PROGRAM prg_TriBlender
VAR
	enumCurrentState	: ENUM_CurrentState;
	FB_SetProductionParams:FB_SetProductionParams;
//stTriBlender		: ST_TriBlender;
	
	sStateDescription		: STRING;
	sStateInstructions		: STRING;
	iCirculationTimeLeft	: UINT;
	bContinue				: BOOL;
	iCurrentMixingComponent	: INT;
	
	tonStageCirculation		: TON;
	
	///For Visu
	bDisableTime			: BOOL;
	bDisableAmount			: BOOL;
	bDisableName			: BOOL;
	bDisableButton			: BOOL;
	wButtonColor			: DWORD;
	
	trig_JumpToCirScreen	: R_TRIG;

	i						: INT;
	bTesting: BOOL;
END_VAR
VAR_IN_OUT
	stTriblender			: ST_TriBlender;
	fb_TriBlenderPump		: FB_Pump;
END_VAR
VAR_INPUT
	arrComponents	: ARRAY [0..g_Prod.cMaxCompInProduct-1] OF ST_Component;
END_VAR

trig_JumpToCirScreen(CLK:= stTriblender.bStartDisolving);

IF trig_JumpToCirScreen.Q THEN
	VisuElems.CurrentVisu:= 'Main';	
END_IF

Init_act_MixingStates();

stTriblender.bPumpOnFdbk:= fb_TriBlenderPump.bRun;

FB_SetProductionParams(stProdParams:=g_Data.arr_ProdTank[0],bTankInProduction:=bTesting,iActualWaterAmount:=100,stTriBlender:=g_Data.stTriBlender);

ACTION CheckIfLast_entry:
bDisableButton:=FALSE;

fb_TriBlenderPump.m_Stop();
bContinue:=FALSE;
END_ACTION

ACTION FlowOrPressureError_entry:
stTriblender.bError:=TRUE;
stTriblender.sErrorDescription:='Pressure or flow error';
VisuElems.CurrentVisu:= 'StartVisu';
END_ACTION

ACTION Init_act_MixingStates:
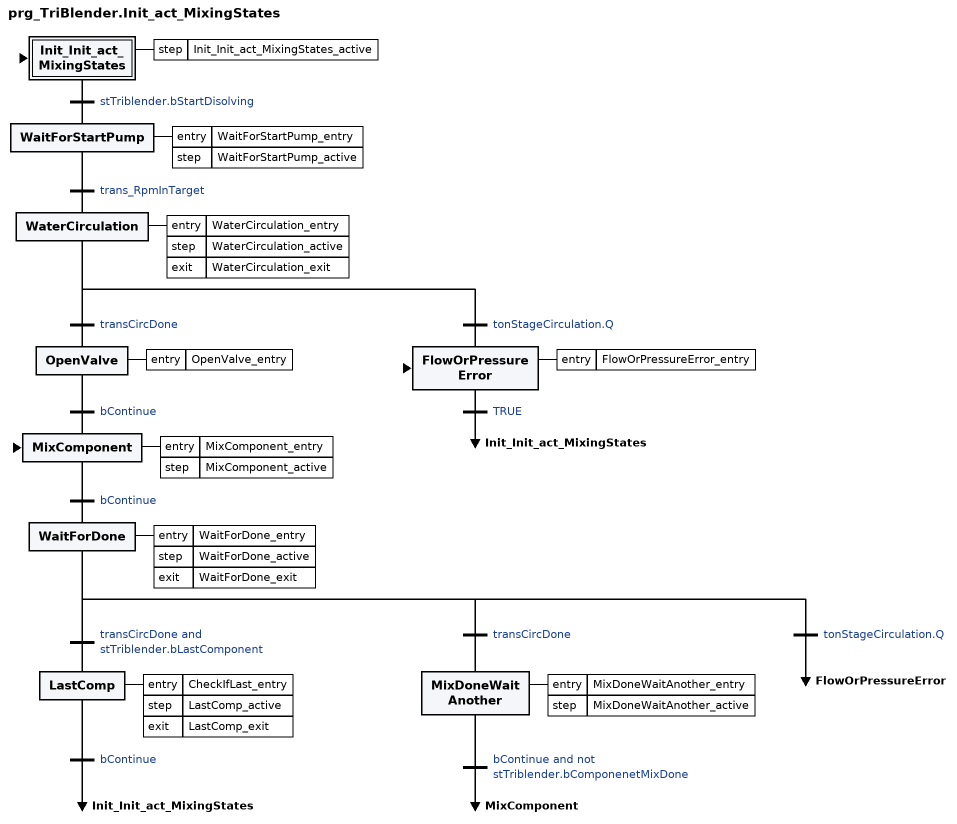
INITIAL_STEP Init_Init_act_MixingStates:
    Init_Init_act_MixingStates_active(N);  // step action
END_STEP
TRANSITION FROM Init_Init_act_MixingStates TO WaitForStartPump
    := stTriblender.bStartDisolving;
END_TRANSITION
STEP WaitForStartPump:
    WaitForStartPump_entry(P1);  // entry action
    WaitForStartPump_active(N);  // step action
END_STEP
TRANSITION FROM WaitForStartPump TO WaterCirculation
    := trans_RpmInTarget;
END_TRANSITION
STEP WaterCirculation:
    WaterCirculation_entry(P1);  // entry action
    WaterCirculation_active(N);  // step action
    WaterCirculation_exit(P0);  // exit action
END_STEP
TRANSITION FROM WaterCirculation TO OpenValve
    := transCircDone;
END_TRANSITION
TRANSITION FROM WaterCirculation TO FlowOrPressureError
    := tonStageCirculation.Q;
END_TRANSITION
STEP FlowOrPressureError:
    FlowOrPressureError_entry(P1);  // entry action
END_STEP
TRANSITION FROM FlowOrPressureError TO Init_Init_act_MixingStates
    := TRUE;
END_TRANSITION
STEP OpenValve:
    OpenValve_entry(P1);  // entry action
END_STEP
TRANSITION FROM OpenValve TO MixComponent
    := bContinue;
END_TRANSITION
STEP MixComponent:
    MixComponent_entry(P1);  // entry action
    MixComponent_active(N);  // step action
END_STEP
TRANSITION FROM MixComponent TO WaitForDone
    := bContinue;
END_TRANSITION
STEP WaitForDone:
    WaitForDone_entry(P1);  // entry action
    WaitForDone_active(N);  // step action
    WaitForDone_exit(P0);  // exit action
END_STEP
TRANSITION FROM WaitForDone TO LastComp
    := transCircDone and stTriblender.bLastComponent;
END_TRANSITION
TRANSITION FROM WaitForDone TO MixDoneWaitAnother
    := transCircDone;
END_TRANSITION
TRANSITION FROM WaitForDone TO FlowOrPressureError
    := tonStageCirculation.Q;
END_TRANSITION
STEP MixDoneWaitAnother:
    MixDoneWaitAnother_entry(P1);  // entry action
    MixDoneWaitAnother_active(N);  // step action
END_STEP
TRANSITION FROM MixDoneWaitAnother TO MixComponent
    := bContinue and not stTriblender.bComponenetMixDone;
END_TRANSITION
STEP LastComp:
    CheckIfLast_entry(P1);  // entry action
    LastComp_active(N);  // step action
    LastComp_exit(P0);  // exit action
END_STEP
TRANSITION FROM LastComp TO Init_Init_act_MixingStates
    := bContinue;
END_TRANSITION
// branch label Branch1_Init_act_MixingStates
// branch label Branch2_Init_act_MixingStates
// branch label Branch0_Init_act_MixingStates
END_ACTION

ACTION Init_Init_act_MixingStates_active:
sStateDescription	:='Triblender valve closed';
sStateInstructions	:= 'Close triblender valve';

bDisableAmount:=TRUE;
bDisableName:=TRUE;
bDisableTime:=TRUE;

wButtonColor:=16#FFC0C0C0;
stTriblender.bError:=FALSE;
stTriblender.bDisolvingDone:=FALSE;
END_ACTION

ACTION LastComp_active:
wButtonColor:=16#FF00FFFF;

sStateDescription	:=	'Finish';
sStateInstructions	:= 	'LastComponentMixed';

bDisableAmount	:=FALSE;
bDisableName	:=FALSE;
bDisableTime	:=FALSE;
END_ACTION

ACTION LastComp_exit:
VisuElems.CurrentVisu:= 'StartVisu';
stTriblender.bDisolvingDone:=TRUE;
END_ACTION

ACTION MixComponent_active:
sStateDescription	:=	'Component Inside';
sStateInstructions	:= 	'Insert component in
 the specified amount';
END_ACTION

ACTION MixComponent_entry:
bContinue:=FALSE;

bDisableAmount	:=FALSE;
bDisableName	:=FALSE;
bDisableTime	:=FALSE;

wButtonColor:=16#FFFF0000;
IF iCurrentMixingComponent<g_Prod.cMaxCompInProduct-1 THEN
	stTriblender.bLastComponent:=NOT arrComponents[iCurrentMixingComponent+1].bComponentEnable;
END_IF
stTriblender.sComponenetAmount:=TO_STRING(arrComponents[iCurrentMixingComponent].rCompActWeight);
stTriblender.sComponenetName:=arrComponents[iCurrentMixingComponent].sDescription;
stTriblender.tComponenetMixingTime:=TO_TIME(arrComponents[iCurrentMixingComponent].iMixingTime*1000);
fb_TriBlenderPump.m_Run(RPM:=arrComponents[iCurrentMixingComponent].rRpmTarget);
END_ACTION

ACTION MixDoneWaitAnother_active:
sStateDescription	:='Triblender valve Opened';
sStateInstructions	:= 'Mix Component done,
 open triblender valve';
END_ACTION

ACTION MixDoneWaitAnother_entry:
bContinue:=FALSE;

bDisableAmount:=TRUE;
bDisableName:=TRUE;
bDisableTime:=TRUE;
bDisableButton:=FALSE;
VisuElems.CurrentVisu:= 'StartVisu';



wButtonColor:=16#FF00FF00;
END_ACTION

ACTION OpenValve_entry:
bContinue:=FALSE;

bDisableAmount:=TRUE;
bDisableName:=TRUE;
bDisableTime:=TRUE;
bDisableButton:=FALSE;

tonStageCirculation(IN:=FALSE);


sStateDescription	:='Triblender valve Opened';
sStateInstructions	:= 'Open triblender valve';

wButtonColor:=16#FF00FF00;
END_ACTION

TRANSITION trans_RpmInTarget:
fb_TriBlenderPump.nRPM< arrComponents[i].rRpmTarget+10 and fb_TriBlenderPump.nRPM> arrComponents[i].rRpmTarget-10
END_TRANSITION

TRANSITION transCircDone:
tonStageCirculation.Q and stTriblender.rMaxAllowedPressure> stTriblender.rPressure and stTriblender.rMinAllowedFlow< stTriblender.rFlow
END_TRANSITION

ACTION WaitForDone_active:
tonStageCirculation(IN:= TRUE,PT:=stTriblender.tComponenetMixingTime);
iCirculationTimeLeft:= TO_UINT(tonStageCirculation.PT - tonStageCirculation.ET)/1000;
bDisableButton:=TRUE;
END_ACTION

ACTION WaitForDone_entry:
wButtonColor:=16#FF0000FF;

sStateDescription	:=	'Waiting';
sStateInstructions	:= 	'Wait for mixing done';
bContinue:=FALSE;

bDisableAmount	:=FALSE;
bDisableName	:=FALSE;
bDisableTime	:=FALSE;


tonStageCirculation(IN:= FALSE);
END_ACTION

ACTION WaitForDone_exit:
stTriblender.bComponenetMixDone:=TRUE;
wButtonColor:=16#FF00FF00;

bDisableAmount	:=TRUE;
bDisableName	:=TRUE;
bDisableTime	:=TRUE;


tonStageCirculation(IN:= FALSE);
END_ACTION

ACTION WaitForStartPump_active:
sStateDescription	:='Start Water Circulation';
sStateInstructions	:= 'Start water circulation, check for leaks';
iCurrentMixingComponent:=0;
bContinue:=FALSE;
FOR i:= 0 TO g_Prod.cMaxCompInProduct-1 DO
	IF arrComponents[i].bIsWater THEN
		fb_TriBlenderPump.m_Run(RPM:=arrComponents[i].rRpmTarget);
	END_IF
END_FOR

wButtonColor:=16#FFFF0000;
END_ACTION

ACTION WaitForStartPump_entry:

stTriblender.bStartDisolving:=FALSE;
END_ACTION

ACTION WaterCirculation_active:
tonStageCirculation(IN:= stTriblender.bPumpOnFdbk,PT:=stTriblender.tWaterCirculationTimeout);
iCirculationTimeLeft:= TO_UINT(tonStageCirculation.PT - tonStageCirculation.ET)/1000;

bDisableButton:=TRUE;

sStateDescription	:='Wait for pressure and flow';
sStateInstructions	:= 'Water circulation in progress,
 check for leaks';
END_ACTION

ACTION WaterCirculation_entry:
bContinue:=FALSE;


bDisableAmount:=TRUE;
bDisableName:=TRUE;
bDisableTime:=FALSE;

tonStageCirculation(IN:=FALSE);
END_ACTION

ACTION WaterCirculation_exit:
tonStageCirculation(IN:=FALSE);
END_ACTION

END_PROGRAM

(* stored: Version 1.1.0.1, ProductVersion 3.1.4024.15
   POU prg_TriBlender: Id {9a86bf9e-8eae-4b5d-8890-d8083718f93d}, SpecialFunc None
   Folder Management: Id {c4ddd0e8-5407-4334-a94a-0f41bc69fac1}
   Action CheckIfLast_entry: Id {0ff06adb-60ce-46ea-a8ba-434fa5634d0f}
   Action FlowOrPressureError_entry: Id {35e66287-119c-40cd-b84f-fa3e256df670}
   Action Init_act_MixingStates: Id {1bb08866-a459-47a2-9078-0401e5c0bb96}
   Action Init_Init_act_MixingStates_active: Id {5b96ca2f-dac9-4416-a4c9-760e9f673ad5}
   Action LastComp_active: Id {2582a41b-802e-45c9-b5d0-7d9f66243cf9}
   Action LastComp_exit: Id {adb66592-836d-46a4-a518-d754da30efe6}
   Action MixComponent_active: Id {1cf67d45-d09f-49f5-ad87-5f9ec42fdf26}
   Action MixComponent_entry: Id {741dfb45-7e63-4493-9a19-e4aebedfdc46}
   Action MixDoneWaitAnother_active: Id {7d82f5bc-b6bc-4046-b841-839403eb7c9b}
   Action MixDoneWaitAnother_entry: Id {ef359ffe-0713-42c1-bf19-c582d7c20eb8}
   Action OpenValve_entry: Id {0d91f935-6559-426a-8a27-b3291b9477d1}
   Transition trans_RpmInTarget: Id {9c69763e-6f57-4306-994c-85c1a23b4746}
   Transition transCircDone: Id {c004dd09-02f8-4be2-a090-e7d683131b10}
   Action WaitForDone_active: Id {b01908cf-9a52-4e61-956b-d173f0b8e957}
   Action WaitForDone_entry: Id {a6f41bb9-a823-4292-995c-7ece526c63aa}
   Action WaitForDone_exit: Id {987162f7-5bc5-4025-8270-3ef2e2dd7475}
   Action WaitForStartPump_active: Id {ede2e026-6ebe-4290-b268-7d5f0ce1e1d3}
   Action WaitForStartPump_entry: Id {59115d06-ebf0-45e1-9214-3f31cd33f08b}
   Action WaterCirculation_active: Id {4f4fcdfa-6e26-4f6f-8974-552317f91ea0}
   Action WaterCirculation_entry: Id {a6b6879f-7055-4ce7-8b92-baa3c44e6dec}
   Action WaterCirculation_exit: Id {a38de536-3fb4-4fcb-9003-5477db64c93a} *)
